// TIA Portal project "040_s71200" (V21)

(* hardware
DEVICE "PLC_1"  S7-1200 Station
   slot 0: "Rack_0"  S7-1200 Rack  Rack  V1.0
   slot 1: "PLC_1"  CPU 1214C DC/DC/DC  6ES7 214-1AG40-0XB0  V4.7
*)

// ===== PLC "PLC_1"  CPU 1214C DC/DC/DC =====

FUNCTION_BLOCK "FB_Lad_ex134"   // FB1, LAD
{ S7_Optimized_Access := 'TRUE' }
   VAR_INPUT
      v_pwm : Hw_Pwm;
      v_enable : Bool;
   END_VAR
   VAR_OUTPUT
      v_busy : Bool;
      v_status : Word;
   END_VAR
   VAR
      inst : CTRL_PWM;
   END_VAR
BEGIN

REGION Network 1: CTRL_PWM - Pulse-width modulation
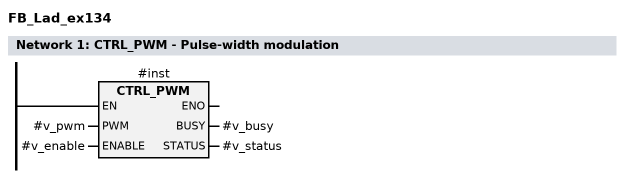
   #inst(PWM := #v_pwm, ENABLE := #v_enable, BUSY => #v_busy, STATUS => #v_status);   // CTRL_PWM
END_REGION
END_FUNCTION_BLOCK

FUNCTION_BLOCK "FB_Fbd_ex134"   // FB2, FBD
{ S7_Optimized_Access := 'TRUE' }
   VAR_INPUT
      v_pwm : Hw_Pwm;
      v_enable : Bool;
   END_VAR
   VAR_OUTPUT
      v_busy : Bool;
      v_status : Word;
   END_VAR
   VAR
      inst : CTRL_PWM;
   END_VAR
BEGIN

REGION Network 1: CTRL_PWM - Pulse-width modulation
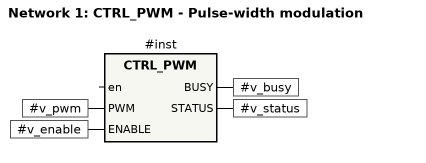
   #inst(PWM := #v_pwm, ENABLE := #v_enable, BUSY => #v_busy, STATUS => #v_status);   // CTRL_PWM
END_REGION
END_FUNCTION_BLOCK

ORGANIZATION_BLOCK "Main"   // OB1, LAD, ProgramCycle
TITLE = "Main Program Sweep (Cycle)"
{ S7_Optimized_Access := 'TRUE' }
VERSION : 0.1
   VAR_INPUT
      Initial_Call : Bool;   // Initial call of this OB
      Remanence : Bool;   // =True, if remanent data are available
   END_VAR
BEGIN
END_ORGANIZATION_BLOCK